Fanuc KAREL source: kb00090.compact.KL

PROGRAM KB00090
%STACKSIZE=65535
%PRIORITY=65535
%NOLOCKGROUP
%ENVIRONMENT REGOPE
VAR
P1 : INTEGER
P2 : BOOLEAN
P3 : INTEGER
P4 : REAL
P5 : INTEGER
BEGIN
P1=1
P2=TRUE
P3=1
P4=1.0
P5=1
GET_REG(P1,P2,P3,P4,P5)
END KB00090
